(* PLC project station_cds.project, CODESYS CODESYS V3.5 SP22 Patch 1 *)
(* stored: creationDateTime 2026-11-25T17:27:32.5174703, modificationDateTime 2026-11-25T17:27:31.3827148 *)

(* Port of OB1 "Main" with the instance DB "InstTestBench": runs the bench by itself after the start. *)
PROGRAM PLC_PRG
  VAR
    Bench : FB_TestBench;
  END_VAR

            Bench();

          
END_PROGRAM
